Fanuc KAREL source: kd00049.KL

PROGRAM KD00049
%STACKSIZE=65535
%PRIORITY=65535
%NOLOCKGROUP
VAR
I : INTEGER
J : INTEGER
B : BOOLEAN
R : REAL
S : STRING[80]
BEGIN
-- UNRESOLVED_PC line 11 opcodes [01 2E 0A 82 0B] marker_code=0
END KD00049
